PROGRAM MAIN
VAR
	tDelayStart : TON;
END_VAR

END_PROGRAM

(* stored: Version 1.1.0.1, ProductVersion 3.1.4024.6
   POU MAIN: Id {883c1222-2c51-4054-8c59-c90c56bed794}, SpecialFunc None *)
